(* IEC 61131-3 sources: StewartPlatform/Network, 1 file *)

(* ---- ConfigObjects.st ---- *)
FUNCTION GLOBAL TAB TASK_CONF
_K_TASK, _K_REAL,
_K_END_VAR,

_K_TASK, _K_CYCLIC,
_K_END_VAR,

_K_TASK, _K_BACKGROUND,
_K_END_VAR,

_K_END_CONF
END_FUNCTION

FUNCTION GLOBAL TAB IPR_CONF
_K_IPR
	0$UINT,
_K_END_VAR,
_K_END_CONF
END_FUNCTION

FUNCTION GLOBAL TAB CONFIG_TABLES
00043$UINT,
0$UINT, 1, 18, "_FILESYS",
0$UINT, 1, 1, "_MULTITASK",
0$UINT, 0, 4, "_OSKERNEL",
0$UINT, 0, 0, "_STDLIB",
0$UINT, 1, 1, "_TASKOBJECTCONTROL",
0$UINT, 1, 30, "AM441",
0$UINT, 1, 18, "BUSINTERFACESDIAS",
0$UINT, 1, 27, "BUSINTERFACESDIASINTERNAL",
0$UINT, 2, 32, "DIASMASTER",
0$UINT, 1, 77, "DIASMASTERC",
0$UINT, 2, 17, "DIASMASTERMAIN",
0$UINT, 1, 0, "DIASMASTERPOSTSCAN",
0$UINT, 1, 9, "DM161",
0$UINT, 1, 11, "EEPROM",
0$UINT, 1, 20, "HUB_BASE",
0$UINT, 2, 10, "HUB_BASE_ROOT",
0$UINT, 2, 32, "HWBASE",
0$UINT, 2, 52, "HWBASECDIAS",
0$UINT, 4, 2, "HWCONTROL",
0$UINT, 1, 10, "HWCONTROLBASE",
0$UINT, 1, 0, "HWRTPOSTSCAN",
0$UINT, 1, 6, "I2CCDIAS",
0$UINT, 0, 0, "IONET",
0$UINT, 1, 21, "MERKEREX",
0$UINT, 1, 9, "RAMFILE",
0$UINT, 1, 3, "SAFETYBASEFSOE",
0$UINT, 3, 8, "SAFETYCDIAS_BASE",
0$UINT, 2, 2, "SAFETYMANAGER",
0$UINT, 1, 10, "SCP111",
0$UINT, 1, 52, "SDIASBASE",
0$UINT, 1, 10, "SDIASHUBBASE",
0$UINT, 1, 81, "SDIASMANAGER",
0$UINT, 1, 44, "SDIASPLC",
0$UINT, 1, 5, "SDIASSAFETYMANAGERFSOE",
0$UINT, 1, 10, "STRING",
0$UINT, 1, 81, "STRINGINTERNAL",
0$UINT, 1, 21, "SYNCCALL",
0$UINT, 2, 9, "VARAN_BASE",
0$UINT, 2, 27, "VARANMANAGER",
0$UINT, 1, 21, "VARANMANAGER_BASE",
0$UINT, 1, 1, "VARANMANAGERPOSTSCAN",
0$UINT, 1, 3, "VIRTUALBASEINIT",
0$UINT, 2, 11, "WATCHDOGDIAS",
ONE_CFG$UINT, 0, 0, "ONE_HW_Network",
ONE_CFG$UINT, 0, 0, "ONE_IONetwork",
TASK_CFG$UINT, 0, 0, "TASK_CONF",
IPR_CFG$UINT, 0, 0, "IPR_CONF",
PRJ_CFG$UINT, 0, 0, "StewartPlatform",
END_FUNCTION

#ifdef __LSLLDR_IOELEMENTS__
FUNCTION GLOBAL TAB _IO_ELEMENTS_TAB
0001$UINT, 0025$UINT,
"Enable_circuit", "DM1611.Output1",
"External_controller", "DM1611.Input6",
"I1", "AM4411.AI1",
"I2", "AM4411.AI2",
"I3", "AM4411.AI3",
"I4", "AM4411.AI4",
"I5", "AM4412.AI1",
"I6", "AM4412.AI2",
"O1", "AM4411.AO1",
"O2", "AM4411.AO2",
"O3", "AM4411.AO3",
"O4", "AM4411.AO4",
"O5", "AM4412.AO1",
"O6", "AM4412.AO2",
"Pressurize", "DM1611.Output4",
"Reset_button", "DM1611.Input5",
"Reset_button_lamp", "DM1611.Output8",
"Reset_EStop", "DM1611.Output5",
"Start_button", "DM1611.Input3",
"Start_button_lamp", "DM1611.Output6",
"Start_pumps", "DM1611.Output3",
"Stop_button", "DM1611.Input4",
"Stop_button_lamp", "DM1611.Output7",
"System_enable_input", "DM1611.Input1",
"System_OK_lamp", "DM1611.Output2",
0025$UINT,
"Enable_circuit", "IONet1.EnableCircuit",
"External_controller", "IONet1.ExternalController",
"I1", "IONet1.I1",
"I2", "IONet1.I2",
"I3", "IONet1.I3",
"I4", "IONet1.I4",
"I5", "IONet1.I5",
"I6", "IONet1.I6",
"O1", "IONet1.O1",
"O2", "IONet1.O2",
"O3", "IONet1.O3",
"O4", "IONet1.O4",
"O5", "IONet1.O5",
"O6", "IONet1.O6",
"Pressurize", "IONet1.Pressurize",
"Reset_button", "IONet1.ResetButton",
"Reset_button_lamp", "IONet1.ResetButtonLamp",
"Reset_EStop", "IONet1.ResetEStop",
"Start_button", "IONet1.StartButton",
"Start_button_lamp", "IONet1.StartButtonLamp",
"Start_pumps", "IONet1.StartPumps",
"Stop_button", "IONet1.StopButton",
"Stop_button_lamp", "IONet1.StopButtonLamp",
"System_enable_input", "IONet1.SystemEnable",
"System_OK_lamp", "IONet1.SystemOKLamp",
END_FUNCTION
#endif //__LSLLDR_IOELEMENTS__
